Universal Robots PolyScope program: restore.urp

Program restore (installation=default_1 directory=/programs/02 Main Routines createdIn=5.19.0 lastSavedIn=5.19.0 robotSerialNumber=20245590068)
Calibrated DH parameters: a=[0.00013, -0.03651, -0.389144, 0.000102, 0.000008, 0]; d=[0.162613, 192.230671, -179.915756, -12.181517, 0.099698, 0.099535]; alpha=[1.57038, 0.002205, 0.004138, 1.570804, -1.571025, 0]; deltaTheta=[-0.000001, 1.484886, 4.928506, -0.130209, 0, 0]
InitVariablesNode
Robot Program (runOnlyOnce=false)
  MoveJ speed 60 deg/s, acceleration 80 deg/s^2 (useActiveTCP=true) feature=Base
    Waypoint Waypoint_1: TCP in base x=2.72 y=-401.535 z=455.349 mm, rx=-3.1317 ry=-0.0062 rz=0.0072 rad; joints [-70.16, -74.711, -107.852, -88.044, 90.079, -160.386] deg; TCP offset x=0 y=0 z=0 mm, rx=0 ry=0 rz=0 rad
